Staubli VAL3: default.pjx

--- default.pjx ---
Parameters millimeterUnit=true stackSize=5000 version=s8.15.1cs9_BS3177
Program file=start.pgx
Program file=stop.pgx
Data file=default.dtx

--- default.dtx ---
mdesc mNomSpeed = {blend=joint, accel=100, vel=100, decel=100, tmax=99999, rmax=99999, leave=50, reach=50}

--- start.pgx ---
program start()
begin
end

--- stop.pgx ---
program stop()
begin
end
